                num nValue[3]
            mdesc mMdesc
            num nActionIndex = 8
            num nDelay
            num nMoveType = 3
            num nPercentage
            num nSigValue = 1
        pointRx pPointRx[2] = {x=594.549819, y=30.770866, z=171.45682, rx=-40.410864, ry=94.502866, rz=40.920287, shoulder=lefty, elbow=epositive, wrist=wnegative}
        string sID
      [76]
        bool bMarked
        jointRx jJointRx = {j1=-1.639134, j2=22.193742, j3=116.03978, j4=1.817031, j5=-44.819098, j6=-0.790246}
        pointRx pInter
        paraItem pParaItem
          [0]
            bool bSafePoint
            ifItem iIfItem
              [0]
                bool bANDOR[2]
                num nSigIndex[3]
                num nSigType[3]
                num nValue[3]
            mdesc mMdesc = {accel=25, vel=50, leave=1}
            num nActionIndex = 8
            num nDelay = 1.8
            num nMoveType = 7
            num nPercentage
            num nSigValue = 1
        pointRx pPointRx[2] = {x=594.549757, y=30.770873, z=70.540177, rx=-40.399083, ry=94.503271, rz=40.908669, shoulder=lefty, elbow=epositive, wrist=wnegative}
        string sID
      [77]
        bool bMarked
        jointRx jJointRx = {j1=-1.639045, j2=12.402747, j3=111.595585, j4=2.517874, j5=-30.594648, j6=-1.669011}
        pointRx pInter
        paraItem pParaItem
          [0]
            bool bSafePoint
            ifItem iIfItem
              [0]
                bool bANDOR[2]
                num nSigIndex[3]
                num nSigType[3]
                num nValue[3]
            mdesc mMdesc
            num nActionIndex = 10
            num nDelay = 5
            num nMoveType = 4
            num nPercentage
            num nSigValue
        pointRx pPointRx[2] = {x=594.549819, y=30.770866, z=171.45682, rx=-40.410864, ry=94.502866, rz=40.920287, shoulder=lefty, elbow=epositive, wrist=wnegative}
        string sID
      [78]
        bool bMarked
        jointRx jJointRx = {j1=-1.639045, j2=12.402747, j3=111.595585, j4=2.517874, j5=-30.594648, j6=-1.669011}
        pointRx pInter
        paraItem pParaItem
          [0]
            bool bSafePoint
            ifItem iIfItem
              [0]
                bool bANDOR[2]
                num nSigIndex[3]
                num nSigType[3]
                num nValue[3]
            mdesc mMdesc
            num nActionIndex = 10
            num nDelay = 0.5
            num nMoveType = 7
            num nPercentage
            num nSigValue
        pointRx pPointRx[2] = {x=594.549819, y=30.770866, z=171.45682, rx=-40.410864, ry=94.502866, rz=40.920287, shoulder=lefty, elbow=epositive, wrist=wnegative}
        string sID
      [79]
        bool bMarked
        jointRx jJointRx = {j1=-1.639045, j2=12.402747, j3=111.595585, j4=2.517874, j5=-30.594648, j6=-1.669011}
        pointRx pInter
        paraItem pParaItem
          [0]
            bool bSafePoint
            ifItem iIfItem
              [0]
                bool bANDOR[2]
                num nSigIndex[3]
                num nSigType[3]
                num nValue[3]
            mdesc mMdesc
            num nActionIndex = 9
            num nDelay = 5
            num nMoveType = 3
            num nPercentage
            num nSigValue = 1
        pointRx pPointRx[2] = {x=594.549819, y=30.770866, z=171.45682, rx=-40.410864, ry=94.502866, rz=40.920287, shoulder=lefty, elbow=epositive, wrist=wnegative}
        string sID
      [80]
        bool bMarked
        jointRx jJointRx = {j1=-0.679346, j2=15.693333, j3=118.292678, j4=-0.521378, j5=-66.0452778, j6=1.744346}
        pointRx pInter
        paraItem pParaItem
          [0]
            bool bSafePoint
            ifItem iIfItem
              [0]
                bool bANDOR[2]
                num nSigIndex[3]
                num nSigType[3]
                num nValue[3]
            mdesc mMdesc
            num nActionIndex = 9
            num nDelay = 5
            num nMoveType
            num nPercentage
            num nSigValue = 1
        pointRx pPointRx[2] = {x=563.98911, y=44.147723, z=151.556034, rx=0.407814, ry=67.941829, rz=0.899564, shoulder=lefty, elbow=epositive, wrist=wnegative}
        string sID
      [81]
        bool bMarked
        jointRx jJointRx = {j1=-2.687248, j2=16.117165, j3=122.304638, j4=-0.487867, j5=-66.528565, j6=1.978834}
        pointRx pInter
        paraItem pParaItem
          [0]
            bool bSafePoint
            ifItem iIfItem
              [0]
                bool bANDOR[2]
                num nSigIndex[3]
                num nSigType[3]
                num nValue[3]
            mdesc mMdesc
            num nActionIndex = 1
            num nDelay = 5
            num nMoveType = 6
            num nPercentage
            num nSigValue = 1
        pointRx pPointRx[2] = {x=546.855577, y=25.169852, z=121.450925, rx=6.745985, ry=71.76392, rz=-5.460967, shoulder=lefty, elbow=epositive, wrist=wnegative}
        string sID
      [82]
        bool bMarked
        jointRx jJointRx = {j1=-2.687248, j2=16.117165, j3=122.304638, j4=-0.487867, j5=-66.528565, j6=1.978834}
        pointRx pInter
        paraItem pParaItem
          [0]
            bool bSafePoint
            ifItem iIfItem
              [0]
                bool bANDOR[2]
                num nSigIndex[3]
                num nSigType[3]
                num nValue[3]
            mdesc mMdesc
            num nActionIndex = 1
            num nDelay = 5
            num nMoveType = 5
            num nPercentage
            num nSigValue = 1
        pointRx pPointRx[2] = {x=546.855577, y=25.169852, z=121.450925, rx=6.745985, ry=71.76392, rz=-5.460967, shoulder=lefty, elbow=epositive, wrist=wnegative}
        string sID
      [83]
        bool bMarked
        jointRx jJointRx = {j1=-1.639045, j2=12.402747, j3=111.595585, j4=2.517874, j5=-30.594648, j6=-1.669011}
        pointRx pInter
        paraItem pParaItem
          [0]
            bool bSafePoint
            ifItem iIfItem
              [0]
                bool bANDOR[2]
                num nSigIndex[3]
                num nSigType[3]
                num nValue[3]
            mdesc mMdesc
            num nActionIndex = 10
            num nDelay
            num nMoveType = 4
            num nPercentage
            num nSigValue = 1
        pointRx pPointRx[2] = {x=594.549819, y=30.770866, z=171.45682, rx=-40.410864, ry=94.502866, rz=40.920287, shoulder=lefty, elbow=epositive, wrist=wnegative}
        string sID
      [84]
        bool bMarked
        jointRx jJointRx = {j1=-1.639045, j2=12.402747, j3=111.595585, j4=2.517874, j5=-30.594648, j6=-1.669011}
        pointRx pInter
        paraItem pParaItem
          [0]
            bool bSafePoint
            ifItem iIfItem
              [0]
                bool bANDOR[2]
                num nSigIndex[3]
                num nSigType[3]
                num nValue[3]
            mdesc mMdesc
            num nActionIndex = 8
            num nDelay
            num nMoveType = 3
            num nPercentage
            num nSigValue = 1
        pointRx pPointRx[2] = {x=594.549819, y=30.770866, z=171.45682, rx=-40.410864, ry=94.502866, rz=40.920287, shoulder=lefty, elbow=epositive, wrist=wnegative}
        string sID
      [85]
        bool bMarked
        jointRx jJointRx = {j1=-1.639134, j2=22.193742, j3=116.03978, j4=1.817031, j5=-44.819098, j6=-0.790246}
        pointRx pInter
        paraItem pParaItem
          [0]
            bool bSafePoint
            ifItem iIfItem
              [0]
                bool bANDOR[2]
                num nSigIndex[3]
                num nSigType[3]
                num nValue[3]
            mdesc mMdesc = {accel=25, vel=50, leave=1}
            num nActionIndex = 8
            num nDelay = 1.8
            num nMoveType = 7
            num nPercentage
            num nSigValue = 1
        pointRx pPointRx[2] = {x=594.549757, y=30.770873, z=70.540177, rx=-40.399083, ry=94.503271, rz=40.908669, shoulder=lefty, elbow=epositive, wrist=wnegative}
        string sID
      [86]
        bool bMarked
        jointRx jJointRx = {j1=-1.639045, j2=12.402747, j3=111.595585, j4=2.517874, j5=-30.594648, j6=-1.669011}
        pointRx pInter
        paraItem pParaItem
          [0]
            bool bSafePoint
            ifItem iIfItem
              [0]
                bool bANDOR[2]
                num nSigIndex[3]
                num nSigType[3]
                num nValue[3]
            mdesc mMdesc
            num nActionIndex = 10
            num nDelay = 5
            num nMoveType = 4
            num nPercentage
            num nSigValue
        pointRx pPointRx[2] = {x=594.549819, y=30.770866, z=171.45682, rx=-40.410864, ry=94.502866, rz=40.920287, shoulder=lefty, elbow=epositive, wrist=wnegative}
        string sID
      [87]
        bool bMarked
        jointRx jJointRx = {j1=-1.639045, j2=12.402747, j3=111.595585, j4=2.517874, j5=-30.594648, j6=-1.669011}
        pointRx pInter
        paraItem pParaItem
          [0]
            bool bSafePoint
            ifItem iIfItem
              [0]
                bool bANDOR[2]
                num nSigIndex[3]
                num nSigType[3]
                num nValue[3]
            mdesc mMdesc
            num nActionIndex = 10
            num nDelay = 0.8
            num nMoveType = 7
            num nPercentage
            num nSigValue
        pointRx pPointRx[2] = {x=594.549819, y=30.770866, z=171.45682, rx=-40.410864, ry=94.502866, rz=40.920287, shoulder=lefty, elbow=epositive, wrist=wnegative}
        string sID
      [88]
        bool bMarked
        jointRx jJointRx = {j1=-1.639045, j2=12.402747, j3=111.595585, j4=2.517874, j5=-30.594648, j6=-1.669011}
        pointRx pInter
        paraItem pParaItem
          [0]
            bool bSafePoint
            ifItem iIfItem
              [0]
                bool bANDOR[2]
                num nSigIndex[3]
                num nSigType[3]
                num nValue[3]
            mdesc mMdesc
            num nActionIndex = 9
            num nDelay = 5
            num nMoveType = 3
            num nPercentage
            num nSigValue = 1
        pointRx pPointRx[2] = {x=594.549819, y=30.770866, z=171.45682, rx=-40.410864, ry=94.502866, rz=40.920287, shoulder=lefty, elbow=epositive, wrist=wnegative}
        string sID
      [89]
        bool bMarked
        jointRx jJointRx = {j1=-1.639045, j2=12.402747, j3=111.595585, j4=2.517874, j5=-30.594648, j6=-1.669011}
        pointRx pInter
        paraItem pParaItem
          [0]
            bool bSafePoint
            ifItem iIfItem
              [0]
                bool bANDOR[2]
                num nSigIndex[3]
                num nSigType[3]
                num nValue[3]
            mdesc mMdesc
            num nActionIndex = 1
            num nDelay = 5
            num nMoveType = 6
            num nPercentage
            num nSigValue
        pointRx pPointRx[2] = {x=594.549819, y=30.770866, z=171.45682, rx=-40.410864, ry=94.502866, rz=40.920287, shoulder=lefty, elbow=epositive, wrist=wnegative}
        string sID
      [90]
        bool bMarked
        jointRx jJointRx = {j1=-1.639045, j2=12.402747, j3=111.595585, j4=2.517874, j5=-30.594648, j6=-1.669011}
        pointRx pInter
        paraItem pParaItem
          [0]
            bool bSafePoint
            ifItem iIfItem
              [0]
                bool bANDOR[2]
                num nSigIndex[3]
                num nSigType[3]
                num nValue[3]
            mdesc mMdesc
            num nActionIndex = 1
            num nDelay = 5
            num nMoveType = 5
            num nPercentage
            num nSigValue
        pointRx pPointRx[2] = {x=594.549819, y=30.770866, z=171.45682, rx=-40.410864, ry=94.502866, rz=40.920287, shoulder=lefty, elbow=epositive, wrist=wnegative}
        string sID
      [91]
        bool bMarked
        jointRx jJointRx = {j1=-6.648853, j2=-3.725267, j3=129.0447837, j4=-6.346169, j5=-34.648625, j6=4.794531}
        pointRx pInter
        paraItem pParaItem
          [0]
            bool bSafePoint
            ifItem iIfItem
              [0]
                bool bANDOR[2]
                num nSigIndex[3]
                num nSigType[3]
                num nValue[3]
            mdesc mMdesc
            num nActionIndex = 1
            num nDelay = 5
            num nMoveType
            num nPercentage
            num nSigValue
        pointRx pPointRx[2] = {x=472.316116, y=1.608512, z=176.939208, rx=-74.680718, ry=93.157376, rz=74.322316, shoulder=lefty, elbow=epositive, wrist=wnegative}
        string sID
      [92]
        bool bMarked
        jointRx jJointRx = {j1=-1.639045, j2=12.402747, j3=111.595585, j4=2.517874, j5=-30.594648, j6=-1.669011}
        pointRx pInter
        paraItem pParaItem
          [0]
            bool bSafePoint
            ifItem iIfItem
              [0]
                bool bANDOR[2]
                num nSigIndex[3]
                num nSigType[3]
                num nValue[3]
            mdesc mMdesc
            num nActionIndex = 11
            num nDelay = 5
            num nMoveType = 4
            num nPercentage
            num nSigValue = 1
        pointRx pPointRx[2] = {x=594.549819, y=30.770866, z=171.45682, rx=-40.410864, ry=94.502866, rz=40.920287, shoulder=lefty, elbow=epositive, wrist=wnegative}
        string sID
      [93]
        bool bMarked
        jointRx jJointRx = {j1=-1.639045, j2=12.402747, j3=111.595585, j4=2.517874, j5=-30.594648, j6=-1.669011}
        pointRx pInter
        paraItem pParaItem
          [0]
            bool bSafePoint
            ifItem iIfItem
              [0]
                bool bANDOR[2]
                num nSigIndex[3]
                num nSigType[3]
                num nValue[3]
            mdesc mMdesc
            num nActionIndex = 10
            num nDelay = 5
            num nMoveType = 3
            num nPercentage
            num nSigValue
        pointRx pPointRx[2] = {x=594.549819, y=30.770866, z=171.45682, rx=-40.410864, ry=94.502866, rz=40.920287, shoulder=lefty, elbow=epositive, wrist=wnegative}
        string sID
      [94]
        bool bMarked
        jointRx jJointRx = {j1=-1.639045, j2=12.402747, j3=111.595585, j4=2.517874, j5=-30.594648, j6=-1.669011}
        pointRx pInter
        paraItem pParaItem
          [0]
            bool bSafePoint
            ifItem iIfItem
              [0]
                bool bANDOR[2]
                num nSigIndex[3]
                num nSigType[3]
                num nValue[3]
            mdesc mMdesc
            num nActionIndex = 9
            num nDelay = 5
            num nMoveType = 4
            num nPercentage
            num nSigValue
        pointRx pPointRx[2] = {x=594.549819, y=30.770866, z=171.45682, rx=-40.410864, ry=94.502866, rz=40.920287, shoulder=lefty, elbow=epositive, wrist=wnegative}
        string sID
      [95]
        bool bMarked
        jointRx jJointRx = {j1=-1.639045, j2=12.402747, j3=111.595585, j4=2.517874, j5=-30.594648, j6=-1.669011}
        pointRx pInter
        paraItem pParaItem
          [0]
            bool bSafePoint
            ifItem iIfItem
              [0]
                bool bANDOR[2]
                num nSigIndex[3]
                num nSigType[3]
                num nValue[3]
            mdesc mMdesc
            num nActionIndex = 11
            num nDelay = 5
            num nMoveType = 4
            num nPercentage
            num nSigValue
        pointRx pPointRx[2] = {x=594.549819, y=30.770866, z=171.45682, rx=-40.410864, ry=94.502866, rz=40.920287, shoulder=lefty, elbow=epositive, wrist=wnegative}
        string sID
    string sID
  [05 sls02]
    num nFrameIndex
    num nMoveID
    num nToolIndex
    pointItem pPointItem[88]
      [0]
        bool bMarked
        jointRx jJointRx = {j1=-2.594987, j2=-12.391258, j3=136.392534, j4=0.644488, j5=-30.575639, j6=-0.113504}
        pointRx pInter
        paraItem pParaItem
          [0]
            bool bSafePoint
            ifItem iIfItem
              [0]
                bool bANDOR[2]
                num nSigIndex[3]
                num nSigType[3]
                num nValue[3]
            mdesc mMdesc
            num nActionIndex = 11
            num nDelay
            num nMoveType = 4
            num nPercentage
            num nSigValue
        pointRx pPointRx[2] = {x=412.772469, y=30.77087, z=171.456836, rx=-40.418431, ry=94.503508, rz=40.927655, shoulder=lefty, elbow=epositive, wrist=wnegative}
        string sID
      [1]
        bool bMarked
        jointRx jJointRx = {j1=-2.594987, j2=-12.391258, j3=136.392534, j4=0.644488, j5=-30.575639, j6=-0.113504}
        pointRx pInter
        paraItem pParaItem
          [0]
            bool bSafePoint
            ifItem iIfItem
              [0]
                bool bANDOR[2]
                num nSigIndex[3]
                num nSigType[3]
                num nValue[3]
            mdesc mMdesc
            num nActionIndex = 9
            num nDelay
            num nMoveType = 4
            num nPercentage
            num nSigValue = 1
        pointRx pPointRx[2] = {x=412.772469, y=30.77087, z=171.456836, rx=-40.418431, ry=94.503508, rz=40.927655, shoulder=lefty, elbow=epositive, wrist=wnegative}
        string sID
      [2]
        bool bMarked
        jointRx jJointRx = {j1=-6.648888, j2=-3.725245, j3=129.0447888, j4=-6.34617, j5=-34.648619, j6=4.79455}
        pointRx pInter
        paraItem pParaItem
          [0]
            bool bSafePoint
            ifItem iIfItem
              [0]
                bool bANDOR[2]
                num nSigIndex[3]
                num nSigType[3]
                num nValue[3]
            mdesc mMdesc
            num nActionIndex
            num nDelay
            num nMoveType
            num nPercentage
            num nSigValue
        pointRx pPointRx[2] = {x=472.316162, y=1.608216, z=176.938999, rx=-74.680314, ry=93.157419, rz=74.321932, shoulder=lefty, elbow=epositive, wrist=wnegative}
        string sID
      [3]
        bool bMarked
        jointRx jJointRx = {j1=-6.652767, j2=20.832827, j3=135.880999, j4=-3.946436, j5=-65.929599, j6=1.179192}
        pointRx pInter
        paraItem pParaItem
          [0]
            bool bSafePoint
            ifItem iIfItem
              [0]
                bool bANDOR[2]
                num nSigIndex[3]
                num nSigType[3]
                num nValue[3]
            mdesc mMdesc
            num nActionIndex
            num nDelay
            num nMoveType
            num nPercentage
            num nSigValue
        pointRx pPointRx[2] = {x=472.315383, y=1.575881, z=5.379837, rx=-74.70962, ry=93.161274, rz=74.351748, shoulder=lefty, elbow=epositive, wrist=wnegative}
        string sID
      [4]
        bool bMarked
        jointRx jJointRx = {j1=-4.442138, j2=54.343414, j3=89.442018, j4=-2.776421, j5=-107.251075, j6=3.647952}
        pointRx pInter
        paraItem pParaItem
          [0]
            bool bSafePoint
            ifItem iIfItem
              [0]
                bool bANDOR[2]
                num nSigIndex[3]
                num nSigType[3]
                num nValue[3]
            mdesc mMdesc
            num nActionIndex
            num nDelay
            num nMoveType
            num nPercentage
            num nSigValue
        pointRx pPointRx[2] = {x=707.968492, y=-0.208433, z=-14.867098, rx=-0.00592828, ry=36.598054, rz=0.906579, shoulder=lefty, elbow=epositive, wrist=wnegative}
        string sID
      [5]
        bool bMarked
        jointRx jJointRx = {j1=-1.639045, j2=12.402747, j3=111.595585, j4=2.517874, j5=-30.594648, j6=-1.669011}
        pointRx pInter
        paraItem pParaItem
          [0]
            bool bSafePoint
            ifItem iIfItem
              [0]
                bool bANDOR[2]
                num nSigIndex[3]
                num nSigType[3]
                num nValue[3]
            mdesc mMdesc
            num nActionIndex = 1
            num nDelay
            num nMoveType = 6
            num nPercentage
            num nSigValue = 1
        pointRx pPointRx[2] = {x=594.549819, y=30.770866, z=171.45682, rx=-40.410864, ry=94.502866, rz=40.920287, shoulder=lefty, elbow=epositive, wrist=wnegative}
        string sID
      [6]
        bool bMarked
        jointRx jJointRx = {j1=-1.639045, j2=12.402747, j3=111.595585, j4=2.517874, j5=-30.594648, j6=-1.669011}
        pointRx pInter
        paraItem pParaItem
          [0]
            bool bSafePoint
            ifItem iIfItem
              [0]
                bool bANDOR[2]
                num nSigIndex[3]
                num nSigType[3]
                num nValue[3]
            mdesc mMdesc
            num nActionIndex = 1
            num nDelay
            num nMoveType = 5
            num nPercentage
            num nSigValue = 1
        pointRx pPointRx[2] = {x=594.549819, y=30.770866, z=171.45682, rx=-40.410864, ry=94.502866, rz=40.920287, shoulder=lefty, elbow=epositive, wrist=wnegative}
        string sID
      [7]
        bool bMarked
        jointRx jJointRx = {j1=-1.639045, j2=12.402747, j3=111.595585, j4=2.517874, j5=-30.594648, j6=-1.669011}
        pointRx pInter
        paraItem pParaItem
          [0]
            bool bSafePoint
            ifItem iIfItem
              [0]
                bool bANDOR[2]
                num nSigIndex[3]
                num nSigType[3]
                num nValue[3]
            mdesc mMdesc
            num nActionIndex = 10
            num nDelay
            num nMoveType = 4
            num nPercentage
            num nSigValue = 1
        pointRx pPointRx[2] = {x=594.549819, y=30.770866, z=171.45682, rx=-40.410864, ry=94.502866, rz=40.920287, shoulder=lefty, elbow=epositive, wrist=wnegative}
        string sID
      [8]
        bool bMarked
        jointRx jJointRx = {j1=-1.639045, j2=12.402747, j3=111.595585, j4=2.517874, j5=-30.594648, j6=-1.669011}
        pointRx pInter
        paraItem pParaItem
          [0]
            bool bSafePoint
            ifItem iIfItem
              [0]
                bool bANDOR[2]
                num nSigIndex[3]
                num nSigType[3]
                num nValue[3]
            mdesc mMdesc
            num nActionIndex = 8
            num nDelay
            num nMoveType = 3
            num nPercentage
            num nSigValue = 1
        pointRx pPointRx[2] = {x=594.549819, y=30.770866, z=171.45682, rx=-40.410864, ry=94.502866, rz=40.920287, shoulder=lefty, elbow=epositive, wrist=wnegative}
        string sID
      [9]
        bool bMarked
        jointRx jJointRx = {j1=-1.639045, j2=12.402747, j3=111.595585, j4=2.517874, j5=-30.594648, j6=-1.669011}
        pointRx pInter
        paraItem pParaItem
          [0]
            bool bSafePoint
            ifItem iIfItem
              [0]
                bool bANDOR[2]
                num nSigIndex[3]
                num nSigType[3]
                num nValue[3]
            mdesc mMdesc
            num nActionIndex = 8
            num nDelay = 2
            num nMoveType = 7
            num nPercentage
            num nSigValue = 1
        pointRx pPointRx[2] = {x=594.549819, y=30.770866, z=171.45682, rx=-40.410864, ry=94.502866, rz=40.920287, shoulder=lefty, elbow=epositive, wrist=wnegative}
        string sID
      [10]
        bool bMarked
        jointRx jJointRx = {j1=-1.639045, j2=12.402747, j3=111.595585, j4=2.517874, j5=-30.594648, j6=-1.669011}
        pointRx pInter
        paraItem pParaItem
          [0]
            bool bSafePoint
            ifItem iIfItem
              [0]
                bool bANDOR[2]
                num nSigIndex[3]
                num nSigType[3]
                num nValue[3]
            mdesc mMdesc
            num nActionIndex = 10
            num nDelay = 5
            num nMoveType = 4
            num nPercentage
            num nSigValue
        pointRx pPointRx[2] = {x=594.549819, y=30.770866, z=171.45682, rx=-40.410864, ry=94.502866, rz=40.920287, shoulder=lefty, elbow=epositive, wrist=wnegative}
        string sID
      [11]
        bool bMarked
        jointRx jJointRx = {j1=-1.639045, j2=12.402747, j3=111.595585, j4=2.517874, j5=-30.594648, j6=-1.669011}
        pointRx pInter
        paraItem pParaItem
          [0]
            bool bSafePoint
            ifItem iIfItem
              [0]
                bool bANDOR[2]
                num nSigIndex[3]
                num nSigType[3]
                num nValue[3]
            mdesc mMdesc
            num nActionIndex = 10
            num nDelay = 0.5
            num nMoveType = 7
            num nPercentage
            num nSigValue
        pointRx pPointRx[2] = {x=594.549819, y=30.770866, z=171.45682, rx=-40.410864, ry=94.502866, rz=40.920287, shoulder=lefty, elbow=epositive, wrist=wnegative}
        string sID
      [12]
        bool bMarked
        jointRx jJointRx = {j1=-1.639045, j2=12.402747, j3=111.595585, j4=2.517874, j5=-30.594648, j6=-1.669011}
        pointRx pInter
        paraItem pParaItem
          [0]
            bool bSafePoint
            ifItem iIfItem
              [0]
                bool bANDOR[2]
                num nSigIndex[3]
                num nSigType[3]
                num nValue[3]
            mdesc mMdesc
            num nActionIndex = 9
            num nDelay = 5
            num nMoveType = 3
            num nPercentage
            num nSigValue = 1
        pointRx pPointRx[2] = {x=594.549819, y=30.770866, z=171.45682, rx=-40.410864, ry=94.502866, rz=40.920287, shoulder=lefty, elbow=epositive, wrist=wnegative}
        string sID
      [13]
        bool bMarked
        jointRx jJointRx = {j1=-6.995994, j2=22.295183, j3=133.491067, j4=-6.412947, j5=-89.696299, j6=3.773786}
        pointRx pInter
        paraItem pParaItem
          [0]
            bool bSafePoint
            ifItem iIfItem
              [0]
                bool bANDOR[2]
                num nSigIndex[3]
                num nSigType[3]
                num nValue[3]
            mdesc mMdesc
            num nActionIndex
            num nDelay
            num nMoveType
            num nPercentage
            num nSigValue
        pointRx pPointRx[2] = {x=480.297234, y=2.689037, z=45.892011, rx=-0.0295899, ry=66.250693, rz=0.93735, shoulder=lefty, elbow=epositive, wrist=wnegative}
        string sID
      [14]
        bool bMarked
        jointRx jJointRx = {j1=-3.631024, j2=-1.590232, j3=111.256847, j4=-19.293027, j5=-7.965925, j6=19.0488477}
        pointRx pInter
        paraItem pParaItem
          [0]
            bool bSafePoint
            ifItem iIfItem
              [0]
                bool bANDOR[2]
                num nSigIndex[3]
                num nSigType[3]
                num nValue[3]
            mdesc mMdesc = {leave=1}
            num nActionIndex
            num nDelay
            num nMoveType = 1
            num nPercentage
            num nSigValue
        pointRx pPointRx[2] = {x=538.454635, y=20.519182, z=260.791216, rx=-4.395762, ry=102.166176, rz=4.98921, shoulder=lefty, elbow=epositive, wrist=wnegative}
        string sID
      [15]
        bool bMarked
        jointRx jJointRx = {j1=-2.334364, j2=-5.268397, j3=112.836865, j4=-1.917467, j5=-5.341213, j6=2.362596}
        pointRx pInter
        paraItem pParaItem
          [0]
            bool bSafePoint
            ifItem iIfItem
              [0]
                bool bANDOR[2]
                num nSigIndex[3]
                num nSigType[3]
                num nValue[3]
            mdesc mMdesc = {leave=1}
            num nActionIndex = 1
            num nDelay
            num nMoveType = 6
            num nPercentage
            num nSigValue = 1
        pointRx pPointRx[2] = {x=515.505365, y=29.338734, z=273.736407, rx=-9.827138, ry=102.415174, rz=10.549826, shoulder=lefty, elbow=epositive, wrist=wnegative}
        string sID
      [16]
        bool bMarked
        jointRx jJointRx = {j1=-2.334364, j2=-5.268397, j3=112.836865, j4=-1.917467, j5=-5.341213, j6=2.362596}
        pointRx pInter
        paraItem pParaItem
          [0]
            bool bSafePoint
            ifItem iIfItem
              [0]
                bool bANDOR[2]
                num nSigIndex[3]
                num nSigType[3]
                num nValue[3]
            mdesc mMdesc = {leave=1}
            num nActionIndex = 1
            num nDelay
            num nMoveType = 5
            num nPercentage
            num nSigValue = 1
        pointRx pPointRx[2] = {x=515.505365, y=29.338734, z=273.736407, rx=-9.827138, ry=102.415174, rz=10.549826, shoulder=lefty, elbow=epositive, wrist=wnegative}
        string sID
      [17]
        bool bMarked
        jointRx jJointRx = {j1=-1.639045, j2=12.402747, j3=111.595585, j4=2.517874, j5=-30.594648, j6=-1.669011}
        pointRx pInter
        paraItem pParaItem
          [0]
            bool bSafePoint
            ifItem iIfItem
              [0]
                bool bANDOR[2]
                num nSigIndex[3]
                num nSigType[3]
                num nValue[3]
            mdesc mMdesc
            num nActionIndex = 10
            num nDelay
            num nMoveType = 4
            num nPercentage
            num nSigValue = 1
        pointRx pPointRx[2] = {x=594.549819, y=30.770866, z=171.45682, rx=-40.410864, ry=94.502866, rz=40.920287, shoulder=lefty, elbow=epositive, wrist=wnegative}
        string sID
      [18]
        bool bMarked
        jointRx jJointRx = {j1=-1.639045, j2=12.402747, j3=111.595585, j4=2.517874, j5=-30.594648, j6=-1.669011}
        pointRx pInter
        paraItem pParaItem
          [0]
            bool bSafePoint
            ifItem iIfItem
              [0]
                bool bANDOR[2]
                num nSigIndex[3]
                num nSigType[3]
                num nValue[3]
            mdesc mMdesc
            num nActionIndex = 8
            num nDelay
            num nMoveType = 3
            num nPercentage
            num nSigValue = 1
        pointRx pPointRx[2] = {x=594.549819, y=30.770866, z=171.45682, rx=-40.410864, ry=94.502866, rz=40.920287, shoulder=lefty, elbow=epositive, wrist=wnegative}
        string sID
      [19]
        bool bMarked
        jointRx jJointRx = {j1=-1.639045, j2=12.402747, j3=111.595585, j4=2.517874, j5=-30.594648, j6=-1.669011}
        pointRx pInter
        paraItem pParaItem
          [0]
            bool bSafePoint
            ifItem iIfItem
              [0]
                bool bANDOR[2]
                num nSigIndex[3]
                num nSigType[3]
                num nValue[3]
            mdesc mMdesc
            num nActionIndex = 8
            num nDelay = 0.8
            num nMoveType = 7
            num nPercentage
            num nSigValue = 1
        pointRx pPointRx[2] = {x=594.549819, y=30.770866, z=171.45682, rx=-40.410864, ry=94.502866, rz=40.920287, shoulder=lefty, elbow=epositive, wrist=wnegative}
        string sID
      [20]
        bool bMarked
        jointRx jJointRx = {j1=-1.639045, j2=12.402747, j3=111.595585, j4=2.517874, j5=-30.594648, j6=-1.669011}
        pointRx pInter
        paraItem pParaItem
          [0]
            bool bSafePoint
            ifItem iIfItem
              [0]
                bool bANDOR[2]
                num nSigIndex[3]
                num nSigType[3]
                num nValue[3]
            mdesc mMdesc
            num nActionIndex = 10
            num nDelay = 5
            num nMoveType = 4
            num nPercentage
            num nSigValue
        pointRx pPointRx[2] = {x=594.549819, y=30.770866, z=171.45682, rx=-40.410864, ry=94.502866, rz=40.920287, shoulder=lefty, elbow=epositive, wrist=wnegative}
        string sID
      [21]
        bool bMarked
        jointRx jJointRx = {j1=-1.639045, j2=12.402747, j3=111.595585, j4=2.517874, j5=-30.594648, j6=-1.669011}
        pointRx pInter
        paraItem pParaItem
          [0]
            bool bSafePoint
            ifItem iIfItem
              [0]
                bool bANDOR[2]
                num nSigIndex[3]
                num nSigType[3]
                num nValue[3]
            mdesc mMdesc
            num nActionIndex = 10
            num nDelay = 0.5
            num nMoveType = 7
            num nPercentage
            num nSigValue
        pointRx pPointRx[2] = {x=594.549819, y=30.770866, z=171.45682, rx=-40.410864, ry=94.502866, rz=40.920287, shoulder=lefty, elbow=epositive, wrist=wnegative}
        string sID
      [22]
        bool bMarked
        jointRx jJointRx = {j1=-1.639045, j2=12.402747, j3=111.595585, j4=2.517874, j5=-30.594648, j6=-1.669011}
        pointRx pInter
        paraItem pParaItem
          [0]
            bool bSafePoint
            ifItem iIfItem
              [0]
                bool bANDOR[2]
                num nSigIndex[3]
                num nSigType[3]
                num nValue[3]
            mdesc mMdesc
            num nActionIndex = 9
            num nDelay = 5
            num nMoveType = 3
            num nPercentage
            num nSigValue = 1
        pointRx pPointRx[2] = {x=594.549819, y=30.770866, z=171.45682, rx=-40.410864, ry=94.502866, rz=40.920287, shoulder=lefty, elbow=epositive, wrist=wnegative}
        string sID
      [23]
        bool bMarked
        jointRx jJointRx = {j1=-4.634649, j2=20.886235, j3=119.504867, j4=-4.475678, j5=-71.496525, j6=3.131235}
        pointRx pInter
        paraItem pParaItem
          [0]
            bool bSafePoint
            ifItem iIfItem
              [0]
                bool bANDOR[2]
                num nSigIndex[3]
                num nSigType[3]
                num nValue[3]
            mdesc mMdesc
            num nActionIndex = 9
            num nDelay = 5
            num nMoveType
            num nPercentage
            num nSigValue = 1
        pointRx pPointRx[2] = {x=568.332279, y=11.51562, z=105.471405, rx=0.230569, ry=69.0075856, rz=-0.170354, shoulder=lefty, elbow=epositive, wrist=wnegative}
        string sID
      [24]
        bool bMarked
        jointRx jJointRx = {j1=-2.687248, j2=16.117165, j3=122.304638, j4=-0.487867, j5=-66.528565, j6=1.978834}
        pointRx pInter
        paraItem pParaItem
          [0]
            bool bSafePoint
            ifItem iIfItem
              [0]
                bool bANDOR[2]
                num nSigIndex[3]
                num nSigType[3]
                num nValue[3]
            mdesc mMdesc
            num nActionIndex = 1
            num nDelay = 5
            num nMoveType = 6
            num nPercentage
            num nSigValue = 1
        pointRx pPointRx[2] = {x=546.855577, y=25.169852, z=121.450925, rx=6.745985, ry=71.76392, rz=-5.460967, shoulder=lefty, elbow=epositive, wrist=wnegative}
        string sID
      [25]
        bool bMarked
        jointRx jJointRx = {j1=-2.687248, j2=16.117165, j3=122.304638, j4=-0.487867, j5=-66.528565, j6=1.978834}
        pointRx pInter
        paraItem pParaItem
          [0]
            bool bSafePoint
            ifItem iIfItem
              [0]
                bool bANDOR[2]
                num nSigIndex[3]
                num nSigType[3]
                num nValue[3]
            mdesc mMdesc
            num nActionIndex = 1
            num nDelay = 5
            num nMoveType = 5
            num nPercentage
            num nSigValue = 1
        pointRx pPointRx[2] = {x=546.855577, y=25.169852, z=121.450925, rx=6.745985, ry=71.76392, rz=-5.460967, shoulder=lefty, elbow=epositive, wrist=wnegative}
        string sID
      [26]
        bool bMarked
        jointRx jJointRx = {j1=-1.639045, j2=12.402747, j3=111.595585, j4=2.517874, j5=-30.594648, j6=-1.669011}
        pointRx pInter
        paraItem pParaItem
          [0]
